FUNCTION_BLOCK DefaultContext EXTENDS TcoCore.TcoContext
VAR
	{attribute addProperty _moveHomeDefaultName "<#MOVE HOME#>"}
	{attribute addProperty _moveWorkDefaultName "<#MOVE TO WORK#>"}
	{attribute addProperty _stopDefaultName "<#STOP a#>"}
    _wpfCyclinder : TcoPneumatics.TcoCylinder(THIS^);
	{attribute addProperty _moveHomeDefaultName "<#MOVE HOME#>"}
	{attribute addProperty _moveWorkDefaultName "<#MOVE TO WORK#>"}
	{attribute addProperty _stopDefaultName "<#STOPDOUBLE#>"}
    _wpfDoubleCyclinder : TcoPneumatics.TcoDoubleCylinder(THIS^);
	{attribute addProperty NameMoveHomeTask "<#In task#>"}
    _wpfCyclinder_1 : TcoPneumatics.TcoCylinder(THIS^);
	{attribute addProperty NameMoveHomeTask "<#In task#>"}
    _wpfCyclinder_2 : TcoPneumatics.TcoCylinder(THIS^);
	{attribute addProperty NameMoveHomeTask "<#In task#>"}
    _wpfCyclinder_3 : TcoPneumatics.TcoCylinder(THIS^);
	disableSignalWork: BOOL;
	disableSignalHome: BOOL;
	suspendSignalWork: BOOL;
	suspendSignalHome: BOOL;
	refilCondition: BOOL;
END_VAR

METHOD PROTECTED  Main
VAR

;
END_VAR
THIS^.RtcSynchronize(TRUE, '', 60);

_wpfCyclinder.Service();	

_wpfCyclinder(inoAtHomePos := IO.A1[0],
	inoAtWorkPos := IO.A1[1],
	inoToHomePos := IO.A2[0],
	inoToWorkPos := IO.A2[1]);
	

	
_wpfCyclinder.AbortMoveHome(disableSignalHome);
_wpfCyclinder.AbortMoveWork(disableSignalWork);

_wpfCyclinder.SuspendMoveHome(suspendSignalHome);
_wpfCyclinder.SuspendMoveWork(suspendSignalWork);

//optional blocking options
//_wpfCyclinder.SuspendMoveWorkInverted(suspendSignalWork);	// is basicaly option how to reproduce exaxt symbol and Not condition
//_wpfCyclinder.SuspendMoveWorkExpression(NOT suspendSignalWork,'Your own msg');	// is basicaly option how to reproduce exaxt symbol and Not condition

_wpfCyclinder.Refill(T#200MS);

_wpfDoubleCyclinder.Service();
_wpfDoubleCyclinder(inoAtHomePos1 := IO.A1[0],
	inoAtHomePos2 := IO.A1[1],
	inoAtWorkPos1 := IO.A1[2],
	inoAtWorkPos2 := IO.A1[3],
	inoToHomePos := IO.A2[3],
	inoToWorkPos := IO.A2[4]);
	
_wpfDoubleCyclinder.AbortMoveHome(disableSignalHome);
_wpfDoubleCyclinder.AbortMoveWork(disableSignalWork);

_wpfDoubleCyclinder.SuspendMoveHome(suspendSignalHome);
_wpfDoubleCyclinder.SuspendMoveWork(suspendSignalWork);

//optional blocking options
//_wpfDoubleCyclinder.SuspendMoveWorkInverted(suspendSignalWork);	// is basicaly option how to reproduce exaxt symbol and Not condition
//_wpfDoubleCyclinder.SuspendMoveWorkExpression(NOT suspendSignalWork,'Your own msg');	// is basicaly option how to reproduce exaxt symbol and Not condition

_wpfDoubleCyclinder.Refill(T#200MS);
END_METHOD

END_FUNCTION_BLOCK

(* stored: Version 1.1.0.1, ProductVersion 3.1.4024.12
   POU DefaultContext: Id {9566aeb0-f006-4c52-ace4-7824786d839b}, SpecialFunc None
   Method Main: Id {f765357f-253d-4bf2-baf0-fad144fcb997} *)
